Fanuc KAREL source: KT00885.KL

PROGRAM KT00885
%NOLOCKGROUP
VAR
  Y1: ARRAY[2] OF BYTE
  Y2: ARRAY[2] OF BYTE
  OUT: REAL
BEGIN
  Y1[1] = 2
  Y2[1] = 3
  Y1[1] = 2
  Y2[1] = 3
  OUT = ATAN2(Y1[1], Y1[1])
END KT00885
